  def create_jig_2(id=0, name="", type=0, capacity=0, jig_offset=p[0,0,0,0,0,0]):
      # iformation about used jigs
      return struct(id=id, name=name, type=type, capacity=capacity, jig_offset=jig_offset)
  end

  JIG2 = create_jig_2()
  JIGs = make_list(0, create_jig_2(), 20)

  JIGs.append(create_jig_2(id=1, name="3FG", type=1, capacity=1, jig_offset=p[0,0,0,0,0,0]))
  JIGs.append(create_jig_2(id=2, name="jig input", type=2, capacity=1, jig_offset=p[0,0,0,0,0,-3.927]))
  JIGs.append(create_jig_2(id=3, name="jig output", type=3, capacity=1, jig_offset=p[0,0,0,0,0,0.78]))
  JIGs.append(create_jig_2(id=6, name="jig bin", type=6, capacity=1, jig_offset=p[0,0,0,0,0,0]))
  JIGs.append(create_jig_2(id=7, name="jig sarstedt racks", type=7, capacity=1, jig_offset=p[0,0,-0.02,0,0,0]))
  JIGs.append(create_jig_2(id=8, name="NoK Bin", type=8, capacity=1, jig_offset=p[0,0,0,0,0,0]))
  JIGs.append(create_jig_2(id=9, name="Pick bott jig", type=9, capacity=1, jig_offset=p[0,0,0,0,0,0]))
  JIGs.append(create_jig_2(id=10, name="Place bott jig", type=10, capacity=1, jig_offset=p[0,0,0,0,0,0]))
  JIGs.append(create_jig_2(id=11, name="bottle shake jig", type=11, capacity=1, jig_offset=p[0,0,0,0,0,0]))
  JIGs.append(create_jig_2(id=12, name="Pick Vial jig", type=12, capacity=1, jig_offset=p[0,0,0,0,0,0]))
  JIGs.append(create_jig_2(id=13, name="Place Vial jig", type=13, capacity=1, jig_offset=p[0,0,0,0,0,0]))
  JIGs.append(create_jig_2(id=14, name="Liquid transfer jig", type=14, capacity=1, jig_offset=p[0,0,0,0,0,0]))
  JIGs.append(create_jig_2(id=15, name="Pick station jig", type=15, capacity=1, jig_offset=p[0,0,0,0,0,0]))
  JIGs.append(create_jig_2(id=16, name="Place station jig", type=16, capacity=1, jig_offset=p[0,0,0,0,0,0]))
  JIGs.append(create_jig_2(id=17, name="Weigh station jig", type=17, capacity=1, jig_offset=p[0,0,0,0,0,0]))
  JIGs.append(create_jig_2(id=18, name="Pick station 1", type=18, capacity=1, jig_offset=p[0,0,0,0,0,0]))
  JIGs.append(create_jig_2(id=19, name="Pick station 2", type=19, capacity=1, jig_offset=p[0,0,0,0,0,0]))
  JIGs.append(create_jig_2(id=20, name="Pick station 3", type=20, capacity=1, jig_offset=p[0,0,0,0,0,0]))
  $ 20 "Script: krish.script"
  def vibration_2():
  	set_analog_out(0,0.4)
  	sleep(0.6)
  	set_analog_out(0,0.0)
  	sleep(0.5)
  end

  def vibration_3():
  	set_analog_out(0,0.4)
  	sleep(0.3)
  	set_analog_out(0,0.0)
  	sleep(0.6)
  end

  def vibration_4():
  	set_analog_out(0,0.4)
  	sleep(0.25)
  	set_analog_out(0, 0.0)
  	sleep(1)
  end

  def vibration_1():
  	set_analog_out(0,0.4)
  	sleep(1)
  	set_analog_out(0,0.0)
  	sleep(0)
  end

  def move_tilt_in_steps(PowA_center, final_pose, steps):
  	i = 0
  	while i <= steps:
  		ratio = i / steps
  		pose_step = p[PowA_center[0] + ratio * (final_pose[0] - PowA_center[0]), PowA_center[1] + ratio * (final_pose[1] -PowA_center[1]),PowA_center[2] + ratio * (final_pose[2] - PowA_center[2]), PowA_center[3] + ratio * (final_pose[3] - PowA_center[3]), PowA_center[4] + ratio * (final_pose[4] - PowA_center[4]), PowA_center[5] + ratio * (final_pose[5] - PowA_center[5])]
  		movej(pose_step, a=1.2, v=0.15)
  		sleep(0.1)
  		i = i+1
  	end
  end

  def tilt_container(angle):
  	P_center = get_actual_tcp_pose()
  	hinge_offset = p[0,0,-0.23,0,0,0]
  	pivot_pose = pose_trans(P_center, hinge_offset)
  	pose_rel = pose_trans(pose_inv(pivot_pose), P_center)
  	angle_mid = (angle/2.0)*3.1416/180
  	angle_end = angle*3.1416/180
  	tilt_mid = p[0,0,0, -angle_mid, 0, 0]
  	tilt_end = p[0,0,0, -angle_end, 0, 0]
  	pose_rel_mid = pose_trans(tilt_mid, pose_rel)
  	pose_rel_end = pose_trans(tilt_end, pose_rel)
  	via_pose = pose_trans(pivot_pose, pose_rel_mid)
  	end_pose = pose_trans(pivot_pose, pose_rel_end)
  	movec(via_pose, end_pose, a=0.05, v=0.01, r=0.001)
  	P_center = get_actual_tcp_pose()
  end

  def scoop_powder(P_center):
  	#scoop_via_offset = p[0.05, 0.025, -0.03,0,0,0]
  	#scoop_end_offset = p[0.10, 0.05, -0.06, 0, 0,0]

  	#scoop_via_pose = pose_trans(scoop_start_pose, scoop_via_offset)
  	#scoop_end_pose = pose_trans(scoop_start_pose, scoop_end_offset)

  	#movel(scoop_start_pose, a=0.3, v=0.1)

  	#movec(scoop_via_pose, scoop_end_pose, a=0.3, v=0.1)

  	approach_offset = p[0.03,0,0.10,0,0,0]
  	scoop_radius = 0.03
  	#scoop_center = p[0, -0.01, 0.02, 0, 0, 1.5708]
  	tilt_down = p[0, 0, 0, -0.2618, 0, 0]
  	#scoop_out = p[0,0,0.10, 0, -0.2618,1.5708]
  	lift_offset = p[0, 0, 0.10, 0, 0, 0]
  	vibration_voltage = 4.0
  	vibration_time = 4.0

  	scoop_entry_pose = pose_trans(P_center, approach_offset)
  	movel(scoop_entry_pose, a=0.05, v=0.05)

  	scoop_start_rel = p[scoop_radius, 0, 0.02, 0, 0, 0]

  	rot_mid = p[0, 0, 0, 0, 0, 0.785]
  	rot_end = p[0, 0, 0, 0, 0, 1.5708]

  	scoop_via_rel = pose_trans(rot_mid, scoop_start_rel)
  	scoop_end_rel = pose_trans(rot_end, scoop_start_rel)

  	scoop_start_pose = pose_trans(P_center, scoop_start_rel)
  	scoop_via_pose = pose_trans(P_center, scoop_via_rel)
  	scoop_end_pose = pose_trans(P_center, scoop_end_rel)

  	movel(scoop_start_pose, a=0.03, v=0.05)

  	movec(scoop_via_pose, scoop_end_pose, a=0.03, v=0.05)

  	#scoop_center_pose = pose_trans(P_center, scoop_center)
  	#movel(scoop_center_pose, a=0.03, v=0.05)

  	tilted_pose = pose_trans(tilt_down, pose_trans(pose_inv(P_center), scoop_end_pose))
  	tilted_pose_in_base = pose_trans(P_center, tilted_pose)

  	movel(tilted_pose_in_base, a=0.03, v=0.05)

  	set_analog_out(0, vibration_voltage)
  	sleep(vibration_time)
  	set_analog_out(0, 0.0)

  	#scoop_out_pose = pose_trans(P_center, scoop_out)
  	#movel(scoop_out_pose, a=0.03, v=0.05)

  	tilt_pose_rel = pose_trans(pose_inv(P_center), tilted_pose_in_base)

  	lifted_pose_rel = pose_trans(lift_offset, tilt_pose_rel)

  	lifted_pose = pose_trans(P_center, lifted_pose_rel)
  	movel(lifted_pose, a=0.03, v=0.05)
  end
  $ 21 "Script: Weight_scale_socket.script"
  def get_weight():
  	socket_open("192.168.12.190", 3002)
  	textmsg("socket opened successfully!")
  	socket_send_string("GET_WEIGHT")
  	sync()
  	sleep(0.5)
  	receiveFromServ = socket_read_ascii_float(6)
  	while (receiveFromServ[0] <1):
  		sleep(0.5)
  		receiveFromServ = socket_read_ascii_float(1)
  		textmsg("retrying read:", receiveFromServ)
  	end
  	textmsg("Received weight:", receiveFromServ[1])
  	socket_close()
  	return receiveFromServ[1]
  end

  def tare_scale():
  	socket_open("192.168.12.190", 3002)
  	socket_send_string("TARE")
  	sleep(0.5)
  	socket_close()
  end

  def zero_scale():
  	socket_open("192.168.12.190", 3002)
  	socket_send_string("ZERO")
  	sleep(0.5)
  	socket_close()
  end
  $ 22 "BeforeStarts"
  $ 23 "uLM"
  $ 24 "CMD_Stop≔ False "
  global CMD_Stop=  False
  $ 25 "CMD_Abort≔ False "
  global CMD_Abort=  False
  $ 26 "CMD_Clear≔ False "
  global CMD_Clear=  False
  $ 27 "STATE≔1"
  global STATE=1
  $ 28 "STATE_Info≔''"
  global STATE_Info=""
  $ 29 "ARM_Referenced≔ False "
  global ARM_Referenced=  False
  $ 30 "zero_ftsensor()"
  zero_ftsensor()
  $ 31 "poses init"
  $ 32 "PSE_A≔p[0,0,0,0,0,0]"
  global PSE_A=p[0,0,0,0,0,0]
  $ 33 "PSE_A_H≔p[0,0,0,0,0,0]"
  global PSE_A_H=p[0,0,0,0,0,0]
  $ 34 "PSE_R≔p[0,0,0,0,0,0]"
  global PSE_R=p[0,0,0,0,0,0]
  $ 35 "PSE_R_H≔p[0,0,0,0,0,0]"
  global PSE_R_H=p[0,0,0,0,0,0]
  $ 36 "PSE_T≔p[0,0,0,0,0,0]"
  global PSE_T=p[0,0,0,0,0,0]
  $ 37 "PSE_T_H≔p[0,0,0,0,0,0]"
  global PSE_T_H=p[0,0,0,0,0,0]
  $ 38 "PSE_C_E≔p[0,0,0,0,0,0]"
  global PSE_C_E=p[0,0,0,0,0,0]
  $ 39 "PSE_C_H≔p[0,0,0,0,0,0]"
  global PSE_C_H=p[0,0,0,0,0,0]
  $ 40 "PSE_C_S≔p[0,0,0,0,0,0]"
  global PSE_C_S=p[0,0,0,0,0,0]
  $ 41 "init_home_by_cartesian_pose(p[0,-0.400,0.300,0,0,0])"
  init_home_by_cartesian_pose(p[0,-0.400,0.300,0,0,0])
  $ 42 "Clearing"
  $ 43 "reset_error()"
  reset_error()
  $ 44 "reset_warning()"
  reset_warning()
  $ 45 "uGo"
  $ 47 "ugo_init( True ,'http://192.168.12.120:10001')"
  ugo_init(  True  ,"http://192.168.12.120:10001")
  $ 48 "ugo_update_outputs()"
  ugo_update_outputs()
  $ 49 "App"
  $ 50 "'ADD APPLICATION SPECIFIC COMMANDS'"
  # 'ADD APPLICATION SPECIFIC COMMANDS'
  $ 51 "Tools"
  $ 52 "OBJ_Picked≔gripper_has_object()"
  global OBJ_Picked=gripper_has_object()
  $ 53 "If OBJ_Picked"
  if (OBJ_Picked):
    # begin: URCap Program Node
    #   Source: Robotiq_Grippers, 1.8.4.4844, Robotiq Inc.
    #   Type: Gripper Activate
    $ 54 "Gripper Activate"

    kill rq_gripper_communication_thread
    rq_gripper_communication_thread_started = False

    rq_init_comm_if_connected(9, "1")
    rq_init_comm_if_connected(2, "2")
    rq_init_comm_if_connected(3, "3")
    rq_init_comm_if_connected(4, "4")
    rq_print_connected_grippers()
    rq_gripper_communication_thread = run rq_gripper_communication()

    while(not rq_gripper_communication_thread_started):
        sync()
    end

    rq_set_max_current_for_all_grippers()

    reset_and_activate = False

    rq_activate_all_grippers(False)
    # end: URCap Program Node
  else:
    $ 55 "Else" "noBreak"
    # begin: URCap Program Node
    #   Source: Robotiq_Grippers, 1.8.4.4844, Robotiq Inc.
    #   Type: Gripper Activate
    $ 56 "Gripper Reset and Activate"

    kill rq_gripper_communication_thread
    rq_gripper_communication_thread_started = False

    rq_init_comm_if_connected(9, "1")
    rq_init_comm_if_connected(2, "2")
    rq_init_comm_if_connected(3, "3")
    rq_init_comm_if_connected(4, "4")
    rq_print_connected_grippers()
    rq_gripper_communication_thread = run rq_gripper_communication()

    while(not rq_gripper_communication_thread_started):
        sync()
    end

    rq_set_max_current_for_all_grippers()

    reset_and_activate = True

    rq_activate_all_grippers(True)
    # end: URCap Program Node
  end
  $ 57 "zero_ftsensor()"
  zero_ftsensor()
  $ 58 "EXTT"
  $ 59 "Set GRP_3F_Enable=Off"
  set_standard_digital_out(4, False)
  $ 60 "Set DO[6]=Off"
  set_standard_digital_out(6, False)
  $ 61 "Set GRP_3F_Decap=Off"
  set_standard_digital_out(3, False)
  $ 62 "Set GRP_3F_Cap=Off"
  set_standard_digital_out(2, False)
  $ 63 "Set GRP_3F_Open=Off"
  set_standard_digital_out(5, False)
  $ 64 "PSE_T≔get_tool_free_pose(dir=[0,0,0.150], move_in_base_frame=True)"
  global PSE_T=get_tool_free_pose(dir=[0,0,0.150], move_in_base_frame=True)
  $ 65 "If is_reachable(Base_const, [PSE_T])"
  if (is_reachable(p[0.0,0.0,0.0,0.0,0.0,0.0], [PSE_T])):
    $ 66 "MoveL"
    $ 67 "PSE_T" "breakAfter"
    movel(PSE_T, a=1.2, v=0.15)
  end
  $ 68 "powder dispensing variable init"
  $ 69 "Start_thread≔ False "
  global Start_thread=  False
  $ 70 "vib_mot_thread≔ False "
  global vib_mot_thread=  False
  $ 71 "kp≔0.00005"
  global kp=0.00005
  $ 72 "ki≔0.0005"
  global ki=0.0005
  $ 73 "kd≔0.002"
  global kd=0.002
  $ 74 "dt≔0.02"
  global dt=0.02
  $ 75 "Integral_error≔0"
  global Integral_error=0
  $ 76 "current_error≔0"
  global current_error=0
  $ 77 "previous_error≔0"
  global previous_error=0
  $ 78 "tilt_increment≔0"
  global tilt_increment=0
  $ 80 "diff≔0"
  global diff=0
  $ 81 "current_pose≔get_actual_tcp_pose()"
  global current_pose= get_actual_tcp_pose ()
  $ 82 "Relative_trans≔p[0.4902, -0.65024, -0.22623, 0.019, -0.263, -5.825]"
  global Relative_trans=p[0.4902, -0.65024, -0.22623, 0.019, -0.263, -5.825]
  $ 83 "ContA_plc_offst≔p[-0.00205, 0.02547, 0.03730, -0.03, -2.183, 6.165]"
  global ContA_plc_offst=p[-0.00205, 0.02547, 0.03730, -0.03, -2.183, 6.165]
  $ 84 "PowA_50_offset≔p[0.21808, -0.19943, 0.06584, 0, 0, 0]"
  global PowA_50_offset=p[0.21808, -0.19943, 0.06584, 0, 0, 0]
  $ 651 "Thread_1"
  thread Thread_1():
    while (True):
      $ 652 "If Start_thread≟ True "
      if (Start_thread ==   True  ):
        $ 653 "Weight_value≔get_weight()"
        global Weight_value=get_weight()
        $ 654 "sync()"
        sync()
      end
    end
  end
  threadId_Thread_1 = run Thread_1()
  $ 655 "Thread_2"
  thread Thread_2():
    while (True):
      $ 656 "Loop vib_mot_thread≟ True "
      thread Thread_while_656():
        while (True):
          $ 657 "diff≔Target_weight-Weight_value"
          global diff=Target_weight-Weight_value
          $ 658 "If diff>0.15"
          global thread_flag_658=0
          thread Thread_if_658():
            $ 660 "Set AO[0]=4.0"
            set_standard_analog_out(0, 0.4)
            thread_flag_658 = 1
          end
          if (diff>0.15):
            global thread_handler_658=run Thread_if_658()
            while (thread_flag_658 == 0):
              if not(diff>0.15):
                kill thread_handler_658
                thread_flag_658 = 2
              else:
                sync()
              end
            end
          else:
            thread_flag_658 = 2
          end
          if (thread_flag_658 == 2):
            $ 661 "ElseIf diff≥0.05 and diff≤0.15"
            global thread_flag_661=0
            thread Thread_if_661():
              $ 662 "vibration_2()"
              vibration_2()
              thread_flag_661 = 1
            end
            if (diff >= 0.05 and diff <= 0.15):
              global thread_handler_661=run Thread_if_661()
              while (thread_flag_661 == 0):
                if not(diff >= 0.05 and diff <= 0.15):
                  kill thread_handler_661
                  thread_flag_661 = 2
                else:
                  sync()
                end
              end
            else:
              thread_flag_661 = 2
            end
            if (thread_flag_661 == 2):
              $ 663 "ElseIf diff≥0.01 and diff<0.05"
              if (diff >= 0.01 and diff<0.05):
                $ 664 "vibration_3()"
                vibration_3()
              else:
                $ 665 "ElseIf diff>0 and diff<0.01"
                if (diff>0 and diff<0.01):
                  $ 666 "vibration_4()"
                  vibration_4()
                else:
                  $ 667 "Else" "noBreak"
                  $ 668 "Set AO[0]=0.0"
                  set_standard_analog_out(0, 0.0)
                end
              end
            end
          end
        end
      end
      if (vib_mot_thread ==   True  ):
        global thread_handler_656=run Thread_while_656()
        while (vib_mot_thread ==   True  ):
          sync()
        end
        kill thread_handler_656
      end
      $ 671 "sync()"
      sync()
    end
  end
  threadId_Thread_2 = run Thread_2()
  while (True):
    $ 85 "Robot Program"
    $ 86 "MAIN"
    $ 87 "command_manager(external_control='uGO', cond_suspend=(ITM_Manipulated and AMR_AtTarget and AMR_Charging and AMR_Battery<40), cond_unsuspend=(AMR_Battery≟60))"
    command_manager(external_control="uGO", cond_suspend=(ITM_Manipulated  and  AMR_AtTarget  and  AMR_Charging  and  AMR_Battery<40), cond_unsuspend=(AMR_Battery == 60))
    $ 88 "log_state(STATE_Info)"
    log_state(STATE_Info)
    $ 89 "Switch STATE"
    switch_1 = STATE
    $ 90 "Case 1"
    if (1 == switch_1):
      $ 91 "Stopping"
      $ 92 "STATE_Info≔'Stopping'"
      global STATE_Info="Stopping"
      $ 93 "end_freedrive_mode()"
      end_freedrive_mode()
      $ 94 "Set"
      set_tcp(p[0.0,0.0,0.161,3.1415,0.0,0.0])
      $ 95 "PSE_T≔get_tool_free_pose(dir=[0,0,0.150], move_in_base_frame=True)"
      global PSE_T=get_tool_free_pose(dir=[0,0,0.150], move_in_base_frame=True)
      $ 96 "If is_reachable(Base_const, [PSE_T])"
      if (is_reachable(p[0.0,0.0,0.0,0.0,0.0,0.0], [PSE_T])):
        $ 97 "MoveL"
        $ 98 "PSE_T" "breakAfter"
        movel(PSE_T, a=1.2, v=0.15)
      end
      $ 99 "do_transition(keep_rxry=OBJ_Picked, r=0)"
      do_transition(keep_rxry=OBJ_Picked, r=0)
      $ 108 "Call Sub_AMR_MiR_V3"
      Sub_AMR_MiR_V3()
      $ 109 "If stopping() and AMR_Done"
      if (stopping()  and  AMR_Done):
        $ 110 "STATE≔2"
        global STATE=2
        $ 111 "ugo_update_outputs()"
        ugo_update_outputs()
      end
    elif (2 == switch_1):
      $ 112 "Case 2"
      $ 113 "Stopped"
      $ 114 "STATE_Info≔'Stopped'"
      global STATE_Info="Stopped"
      $ 115 "Call Sub_AMR_MiR_V3"
      Sub_AMR_MiR_V3()
      $ 116 "If CMD_Reset"
      if (CMD_Reset):
        $ 117 "STATE≔3"
        global STATE=3
        $ 118 "ugo_update_outputs()"
        ugo_update_outputs()
      end
    elif (3 == switch_1):
      $ 119 "Case 3"
      $ 120 " Resetting"
      $ 121 "STATE_Info≔'Resetting'"
      global STATE_Info="Resetting"
      $ 122 "uML"
      $ 123 "reset_error()"
      reset_error()
      $ 124 "reset_warning()"
      reset_warning()
      $ 125 "PROCESS_Step≔0"
      global PROCESS_Step=0
      $ 126 "PROCESS_Info≔''"
      global PROCESS_Info=""
      $ 127 "ARM_Referenced≔ False "
      global ARM_Referenced=  False
      $ 128 "WRK_Done≔ False "
      global WRK_Done=  False
      $ 129 "ITM_Prepared≔ False "
      global ITM_Prepared=  False
      $ 130 "ITM_Manipulated≔ False "
      global ITM_Manipulated=  False
      $ 131 "STP≔0"
      global STP=0
      $ 132 "Action≔0"
      global Action=0
      $ 133 "Action_Info≔''"
      global Action_Info=""
      $ 134 "ITM_ID≔0"
      global ITM_ID=0
      $ 135 "JIG≔0"
      global JIG=0
      $ 136 "JIG_Slot≔0"
      global JIG_Slot=0
      $ 137 "Task_info≔''"
      global Task_info=""
      $ 138 "Set"
      set_tcp(p[0.0,0.0,0.161,3.1415,0.0,0.0])
      $ 139 "App"
      $ 140 "'ADD APPLICATION SPECIFIC COMMANDS'"
      # 'ADD APPLICATION SPECIFIC COMMANDS'
      $ 141 "OBJ_Type≔0"
      global OBJ_Type=0
      $ 142 "OBJ_Nbr≔0"
      global OBJ_Nbr=0
      $ 143 "If CNT_Rack_Output≥50"
      if (CNT_Rack_Output >= 50):
        $ 144 "CNT_Rack_Output≔0"
        global CNT_Rack_Output=0
      end
      $ 145 "TASK≔struct(ID=0, NAVI=struct(target=0, footprint=0, protectiveOff=0, dock=0), WORK=struct(ITM_ID_Src=0, JIG_ID_Src=0, OBJ_Nbr_Src=0, ACT_Src=0, ITM_ID_Tgt=0, JIG_ID_Tgt=0, OBJ_Nbr_Tgt=0, ACT_Tgt=0, OBJ_Type=0))"
      global TASK=struct(ID=0, NAVI=struct(target=0, footprint=0, protectiveOff=0, dock=0), WORK=struct(ITM_ID_Src=0, JIG_ID_Src=0, OBJ_Nbr_Src=0, ACT_Src=0, ITM_ID_Tgt=0, JIG_ID_Tgt=0, OBJ_Nbr_Tgt=0, ACT_Tgt=0, OBJ_Type=0))
      $ 146 "Call Sub_AMR_MiR_V3"
      Sub_AMR_MiR_V3()
      $ 147 "If resetting() and AMR_Done"
      if (resetting()  and  AMR_Done):
        $ 148 "STATE≔4"
        global STATE=4
        $ 149 "ugo_update_outputs()"
        ugo_update_outputs()
      end
    elif (4 == switch_1):
      $ 150 "Case 4"
      $ 151 "Idle"
      $ 152 "STATE_Info≔'Idle'"
      global STATE_Info="Idle"
      $ 153 "If CMD_Start"
      if (CMD_Start):
        $ 154 "STATE≔5"
        global STATE=5
        $ 155 "ugo_update_outputs()"
        ugo_update_outputs()
      end
    elif (5 == switch_1):
      $ 156 "Case 5"
      $ 157 "Starting"
      $ 158 "STATE_Info≔'Starting'"
      global STATE_Info="Starting"
      $ 159 "'ADD COMMANDS WHAT TO START WITH'"
      # 'ADD COMMANDS WHAT TO START WITH'
      $ 160 "Call Sub_AMR_MiR_V3"
      Sub_AMR_MiR_V3()
      $ 161 "get ugo data"
      $ 162 "Assign Tasks"
      $ 163 "TASK.ID = ugo_get_task()"
      TASK.ID = ugo_get_task()
      $ 164 "If TASK.ID≟1"
      if (TASK.ID == 1):
        $ 165 "Task_info≔'Charge'"
        global Task_info="Charge"
        $ 166 "Parameters"
        $ 167 "AMR_PosTarget≔1"
        global AMR_PosTarget=1
      else:
        $ 168 "ElseIf TASK.ID≟9"
        if (TASK.ID == 9):
          $ 169 "'Pick Sarstedt Rack from Variable source'"
          # 'Pick Sarstedt Rack from Variable source'
          $ 170 "Task_info≔'Navigate to Target'"
          global Task_info="Navigate to Target"
          $ 171 "Parameters"
          $ 172 "AMR_PosTarget≔UGO.read_input('00','ITM_ID')"
          global AMR_PosTarget=UGO.read_input("00","ITM_ID")
        else:
          $ 173 "ElseIf TASK.ID≟99"
          if (TASK.ID == 99):
            $ 174 "Task_info≔'Pick rack pipet'"
            global Task_info="Pick rack pipet"
            $ 175 "Parameters"
            $ 176 "ITM_ID≔1"
            global ITM_ID=1
            $ 177 "OBJ_Type≔9"
            global OBJ_Type=9
            $ 178 "JIG≔18"
            global JIG=18
            $ 179 "AMR_PosTarget≔3"
            global AMR_PosTarget=3
          else:
            $ 180 "ElseIf TASK.ID≟98"
            if (TASK.ID == 98):
              $ 181 "Task_info≔'Place rack pipet'"
              global Task_info="Place rack pipet"
              $ 182 "Parameters"
              $ 183 "ITM_ID≔1"
              global ITM_ID=1
              $ 184 "OBJ_Type≔9"
              global OBJ_Type=9
              $ 185 "JIG≔19"
              global JIG=19
              $ 186 "AMR_PosTarget≔2"
              global AMR_PosTarget=2
            else:
              $ 187 "Else" "noBreak"
              $ 188 "set_error(ERROR_WRONG_ORDER)"
              set_error(ERROR_WRONG_ORDER)
            end
          end
        end
      end
      $ 189 "test ugo"
      $ 190 "Wait: 0.2"
      sleep(0.2)
      $ 191 "ugo_update_outputs()"
      ugo_update_outputs()
      $ 192 "If starting() and AMR_Done"
      if (starting()  and  AMR_Done):
        $ 193 "log_message(Task_info, 'New Task: ')"
        log_message(Task_info, "New Task: ")
        $ 194 "log_message(to_str(TASK.ID), 'Task_ID: ')"
        log_message(to_str(TASK.ID), "Task_ID: ")
        $ 195 "do_transition(keep_rxry=OBJ_Picked)"
        do_transition(keep_rxry=OBJ_Picked)
        $ 196 "STATE≔6"
        global STATE=6
        $ 197 "ugo_update_outputs()"
        ugo_update_outputs()
      end
    elif (6 == switch_1):
      $ 198 "Case 6"
      $ 199 "Execute"
      $ 200 "STATE_Info≔'Execute'"
      global STATE_Info="Execute"
      $ 201 "If  not CMD_Hold and not CMD_Suspend"
      global thread_flag_201=0
      thread Thread_if_201():
        $ 202 "Switch PROCESS_Step"
        switch_2 = PROCESS_Step
        $ 203 "Case 0"
        if (0 == switch_2):
          $ 204 "PROCESS_Info≔'process control'"
          global PROCESS_Info="process control"
          $ 205 "log_process(PROCESS_Info)"
          log_process(PROCESS_Info)
          $ 206 "process control"
          $ 207 "If  not AMR_AtTarget"
          if (  not  AMR_AtTarget):
            $ 208 "PROCESS_Step≔1"
            global PROCESS_Step=1
          else:
            $ 209 "ElseIf (( not ITM_Prepared and  not WRK_Done) or (ITM_Prepared and WRK_Done))"
            if (((  not  ITM_Prepared  and    not  WRK_Done)  or  (ITM_Prepared  and  WRK_Done))):
              $ 210 "PROCESS_Step≔2"
              global PROCESS_Step=2
            else:
              $ 211 "ElseIf  not WRK_Done"
              if (  not  WRK_Done):
                $ 212 "PROCESS_Step≔3"
                global PROCESS_Step=3
              else:
                $ 213 "Else" "noBreak"
                $ 214 "task finished"
                $ 215 "PROCESS_Info≔''"
                global PROCESS_Info=""
                $ 216 "STATE≔7"
                global STATE=7
                $ 217 "ugo_update_outputs()"
                ugo_update_outputs()
              end
            end
          end
        elif (1 == switch_2):
          $ 218 "Case 1"
          $ 219 "navigate"
          $ 220 "'MOVING THE uML'"
          # 'MOVING THE uML'
          $ 221 "PROCESS_Info≔'move to target'"
          global PROCESS_Info="move to target"
          $ 222 "log_process(PROCESS_Info)"
          log_process(PROCESS_Info)
          $ 223 "If TASK.ID≟1"
          if (TASK.ID == 1):
            $ 224 "Action≔51"
            global Action=51
          else:
            $ 225 "Else" "noBreak"
            $ 226 "Action≔52"
            global Action=52
          end
          $ 227 "Call Sub_AMR_MiR_V3"
          Sub_AMR_MiR_V3()
          $ 228 "If AMR_Done"
          if (AMR_Done):
            $ 229 "PROCESS_Step≔0"
            global PROCESS_Step=0
          end
        elif (2 == switch_2):
          $ 230 "Case 2"
          $ 231 "prepare"
          $ 232 "'THINGS THAT HAVE TO BE DONE ONCE IN A SEQUENCE,WORKFLOW'"
          # 'THINGS THAT HAVE TO BE DONE ONCE IN A SEQUENCE,WORKFLOW'
          $ 233 "PROCESS_Info≔'prepare for work'"
          global PROCESS_Info="prepare for work"
          $ 234 "log_process(PROCESS_Info)"
          log_process(PROCESS_Info)
          $ 235 "If TASK.WORK.ITM_ID_Src>1"
          if (TASK.WORK.ITM_ID_Src>1):
            $ 236 "ITM_ID≔TASK.WORK.ITM_ID_Src"
            global ITM_ID=TASK.WORK.ITM_ID_Src
          else:
            $ 237 "ElseIf TASK.WORK.ITM_ID_Tgt>1"
            if (TASK.WORK.ITM_ID_Tgt>1):
              $ 238 "ITM_ID≔TASK.WORK.ITM_ID_Tgt"
              global ITM_ID=TASK.WORK.ITM_ID_Tgt
            end
          end
          $ 239 "If  not ARM_Referenced and (ITM_ID≠0)"
          if (  not  ARM_Referenced  and  (ITM_ID != 0)):
            $ 240 "STP≔1"
            global STP=1
          else:
            $ 241 "ElseIf ARM_Referenced or (ITM_ID≟0)"
            if (ARM_Referenced  or  (ITM_ID == 0)):
              $ 242 "STP≔2"
              global STP=2
            end
          end
          $ 243 "Switch STP"
          switch_3 = STP
          $ 244 "Case 1"
          if (1 == switch_3):
            $ 245 "reference"
            $ 246 "STP_Info≔'reference at target position'"
            global STP_Info="reference at target position"
            $ 247 "log_step(STP_Info)"
            log_step(STP_Info)
            $ 248 "If ITM_ID≟1"
            if (ITM_ID == 1):
              $ 249 "CAM_Done≔ True "
              global CAM_Done=  True
            else:
              $ 250 "Else" "noBreak"
              $ 251 "Action≔131"
              global Action=131
              $ 252 "Call Sub_Vision_V18"
              Sub_Vision_V18()
            end
            $ 254 "If CAM_Done and  not ERROR.FLAG"
            if (CAM_Done  and    not  ERROR.FLAG):
              $ 255 "log_step('ARM referenced')"
              log_step("ARM referenced")
              $ 256 "ARM_Referenced≔ True "
              global ARM_Referenced=  True
            end
          elif (2 == switch_3):
            $ 257 "Case 2"
            $ 258 "manipulate"
            $ 259 "STP_Info≔'manipulate item'"
            global STP_Info="manipulate item"
            $ 260 "log_step(STP_Info)"
            log_step(STP_Info)
            $ 261 "'In case pressing button is needed'"
            # 'In case pressing button is needed'
            $ 262 "If found_in_list(ITM_ID, ITM_ID_List)"
            if (found_in_list(ITM_ID, ITM_ID_List)):
              $ 263 "Switch ITM_ID"
              switch_4 = ITM_ID
              $ 264 "Case 0"
              if (0 == switch_4):
                $ 265 "ITM_Manipulated≔ not ITM_Manipulated"
                global ITM_Manipulated=  not  ITM_Manipulated
              elif (1 == switch_4):
                $ 266 "Case 1"
                $ 267 "ITM_Manipulated≔ not ITM_Manipulated"
                global ITM_Manipulated=  not  ITM_Manipulated
              elif (2 == switch_4):
                $ 268 "Case 2"
              else:
                $ 278 "Default Case"
                $ 279 "ITM_Manipulated≔ not ITM_Manipulated"
                global ITM_Manipulated=  not  ITM_Manipulated
              end
            end
          end
          $ 280 "ITM_Prepared≔(ITM_Manipulated or  not found_in_list(ITM_ID, ITM_ID_List)) and (ARM_Referenced or ITM_ID≟0) and  not WRK_Done"
          global ITM_Prepared=(ITM_Manipulated  or    not  found_in_list(ITM_ID, ITM_ID_List))  and  (ARM_Referenced  or  ITM_ID == 0)  and    not  WRK_Done
          $ 281 "STP≔0"
          global STP=0
          $ 282 "STP_Info≔''"
          global STP_Info=""
          $ 283 "PROCESS_Step≔0"
          global PROCESS_Step=0
        elif (3 == switch_2):
          $ 284 "Case 3"
          $ 285 "work"
          $ 286 "'ADD EVERY MACHINE, OBJECT, STATION TO WORK ON'"
          # 'ADD EVERY MACHINE, OBJECT, STATION TO WORK ON'
          $ 287 "Switch ITM_ID"
          switch_3 = ITM_ID
          $ 288 "Case 1"
          if (1 == switch_3):
            $ 289 "uLM"
            $ 290 "If TASK.ID≟12"
            if (TASK.ID == 12):
              $ 291 "fill racks"
              $ 292 "Action≔151"
              global Action=151
              $ 293 "Call Sub_Vision_V18"
              Sub_Vision_V18()
              $ 294 "If  not ERROR.FLAG"
              if (  not  ERROR.FLAG):
                $ 295 "Actions for the task"
                $ 296 "Action≔1"
                global Action=1
                $ 297 "JIG≔2"
                global JIG=2
                $ 298 "JIG_Slot≔CAM_Result[0]"
                global JIG_Slot=CAM_Result[0]
                $ 299 "OBJ_Nbr≔CAM_Result[0]"
                global OBJ_Nbr=CAM_Result[0]
                $ 300 "OBJ_Type≔2"
                global OBJ_Type=2
                $ 301 "Call Sub_Action_V4"
                Sub_Action_V4()
                $ 302 "If OBJ_Picked"
                if (OBJ_Picked):
                  $ 303 "CAM_Result.remove(0)"
                  CAM_Result.remove(0)
                  $ 304 "PRC_TubCounter≔PRC_TubCounter+1"
                  global PRC_TubCounter=PRC_TubCounter+1
                  $ 305 "If PRC_TubCounter%4≟0"
                  if (PRC_TubCounter%4 == 0):
                    $ 306 "JIG_Slot≔4"
                    global JIG_Slot=4
                  else:
                    $ 307 "Else" "noBreak"
                    $ 308 "JIG_Slot≔PRC_TubCounter%4"
                    global JIG_Slot=PRC_TubCounter%4
                  end
                  $ 309 "OBJ_Nbr≔ceil(PRC_TubCounter/4)"
                  global OBJ_Nbr=ceil(PRC_TubCounter/4)
                  $ 310 "Action≔2"
                  global Action=2
                  $ 311 "JIG≔4"
                  global JIG=4
                  $ 312 "Call Sub_Action_V4"
                  Sub_Action_V4()
                  $ 313 "Action≔151"
                  global Action=151
                  $ 314 "Call Sub_Vision_V18"
                  Sub_Vision_V18()
                end
              end
              $ 315 "If (CAM_Captures≥CAM_PRM_Retries) or (PRC_TubCounter≥32)"
              if ((CAM_Captures >= CAM_PRM_Retries)  or  (PRC_TubCounter >= 32)):
                $ 316 "PROCESS_Step≔0"
                global PROCESS_Step=0
                $ 317 "WRK_Done≔ True "
                global WRK_Done=  True
              end
            else:
              $ 318 "ElseIf TASK.ID≟49"
              if (TASK.ID == 49):
                $ 319 "Pick Powder container"
                $ 320 "Action≔131"
                global Action=131
                $ 321 "Call Sub_Vision_V18"
                Sub_Vision_V18()
                $ 322 "Action≔35"
                global Action=35
                $ 323 "Call Sub_Action_V4"
                Sub_Action_V4()
                $ 324 "PROCESS_Step≔0"
                global PROCESS_Step=0
                $ 325 "WRK_Done≔ True "
                global WRK_Done=  True
              else:
                $ 326 "ElseIf TASK.ID≟50"
                if (TASK.ID == 50):
                  $ 327 "Decap containers"
                  $ 328 "Action≔36"
                  global Action=36
                  $ 329 "Call Sub_Action_V4"
                  Sub_Action_V4()
                  $ 330 "PROCESS_Step≔0"
                  global PROCESS_Step=0
                  $ 331 "WRK_Done≔ True "
                  global WRK_Done=  True
                else:
                  $ 332 "ElseIf TASK.ID≟51"
                  if (TASK.ID == 51):
                    $ 333 "Detect Spatula and transfer powder"
                    $ 334 "Action≔131"
                    global Action=131
                    $ 335 "Call Sub_Vision_V18"
                    Sub_Vision_V18()
                    $ 336 "Action≔37"
                    global Action=37
                    $ 337 "Call Sub_Action_V4"
                    Sub_Action_V4()
                    $ 338 "PROCESS_Step≔0"
                    global PROCESS_Step=0
                    $ 339 "WRK_Done≔ True "
                    global WRK_Done=  True
                  else:
                    $ 340 "ElseIf TASK.ID≟52"
                    if (TASK.ID == 52):
                      $ 341 "Pick PowderA container"
                      $ 342 "Action≔131"
                      global Action=131
                      $ 343 "Call Sub_Vision_V18"
                      Sub_Vision_V18()
                      $ 344 "Action≔38"
                      global Action=38
                      $ 345 "Call Sub_Action_V4"
                      Sub_Action_V4()
                      $ 346 "PROCESS_Step≔0"
                      global PROCESS_Step=0
                      $ 347 "WRK_Done≔ True "
                      global WRK_Done=  True
                    else:
                      $ 348 "ElseIf TASK.ID≟53"
                      if (TASK.ID == 53):
                        $ 349 "Decap containerA"
                        $ 350 "Action≔39"
                        global Action=39
                        $ 351 "Call Sub_Action_V4"
                        Sub_Action_V4()
                        $ 352 "PROCESS_Step≔0"
                        global PROCESS_Step=0
                        $ 353 "WRK_Done≔ True "
                        global WRK_Done=  True
                      else:
                        $ 354 "ElseIf TASK.ID≟54"
                        if (TASK.ID == 54):
                          $ 355 "Dispense PowderA"
                          $ 356 "Action≔131"
                          global Action=131
                          $ 357 "Call Sub_Vision_V18"
                          Sub_Vision_V18()
                          $ 358 "Action≔40"
                          global Action=40
                          $ 359 "Call Sub_Action_V4"
                          Sub_Action_V4()
                          $ 360 "PROCESS_Step≔0"
                          global PROCESS_Step=0
                          $ 361 "WRK_Done≔ True "
                          global WRK_Done=  True
                        else:
                          $ 362 "ElseIf TASK.ID≟54"
                          if (TASK.ID == 54):
                            $ 363 "Dispense PowderA"
                            $ 364 "Action≔131"
                            global Action=131
                            $ 365 "Call Sub_Vision_V18"
                            Sub_Vision_V18()
                            $ 366 "Action≔40"
                            global Action=40
                            $ 367 "Call Sub_Action_V4"
                            Sub_Action_V4()
                            $ 368 "PROCESS_Step≔0"
                            global PROCESS_Step=0
                            $ 369 "WRK_Done≔ True "
                            global WRK_Done=  True
                          else:
                            $ 370 "ElseIf TASK.ID≟99"
                            if (TASK.ID == 99):
                              $ 371 "Pick rack pipet"
                              $ 372 "Action≔131"
                              global Action=131
                              $ 373 "Call Sub_Vision_V18"
                              Sub_Vision_V18()
                              $ 374 "Action≔5"
                              global Action=5
                              $ 375 "Call Sub_Action_V4"
                              Sub_Action_V4()
                              $ 376 "PROCESS_Step≔0"
                              global PROCESS_Step=0
                              $ 377 "WRK_Done≔ True "
                              global WRK_Done=  True
                            else:
                              $ 378 "ElseIf TASK.ID≟98"
                              if (TASK.ID == 98):
                                $ 379 "Pick rack pipet"
                                $ 380 "Action≔131"
                                global Action=131
                                $ 381 "Call Sub_Vision_V18"
                                Sub_Vision_V18()
                                $ 382 "Action≔6"
                                global Action=6
                                $ 383 "Call Sub_Action_V4"
                                Sub_Action_V4()
                                $ 384 "PROCESS_Step≔0"
                                global PROCESS_Step=0
                                $ 385 "WRK_Done≔ True "
                                global WRK_Done=  True
                              end
                            end
                          end
                        end
                      end
                    end
                  end
                end
              end
            end
          elif (2 == switch_3):
            $ 386 "Case 2"
          elif (5 == switch_3):
            $ 428 "Case 5"
          elif (20 == switch_3):
            $ 436 "Case 20"
          elif (43 == switch_3):
            $ 498 "Case 43"
          else:
            $ 506 "Default Case"
            $ 507 "WRK_Done≔ True "
            global WRK_Done=  True
            $ 508 "PROCESS_Step≔0"
            global PROCESS_Step=0
          end
        end
        thread_flag_201 = 1
      end
      if (  not  CMD_Hold and not CMD_Suspend):
        global thread_handler_201=run Thread_if_201()
        while (thread_flag_201 == 0):
          if not(  not  CMD_Hold and not CMD_Suspend):
            kill thread_handler_201
            thread_flag_201 = 2
          else:
            sync()
          end
        end
      else:
        thread_flag_201 = 2
      end
      $ 509 "If CMD_Hold"
      if (CMD_Hold):
        $ 510 "STATE≔9"
        global STATE=9
        $ 511 "ugo_update_outputs()"
        ugo_update_outputs()
      else:
        $ 512 "ElseIf CMD_Suspend"
        if (CMD_Suspend):
          $ 513 "STATE≔12"
          global STATE=12
          $ 514 "ugo_update_outputs()"
          ugo_update_outputs()
        end
      end
    elif (7 == switch_1):
      $ 515 "Case 7"
      $ 516 "Completing"
      $ 517 "STATE_Info≔'Completing'"
      global STATE_Info="Completing"
      $ 518 "'ADD COMMANDS FOR COMPLETING THE PROCESS'"
      # 'ADD COMMANDS FOR COMPLETING THE PROCESS'
      $ 519 "do_transition(keep_rxry=OBJ_Picked)"
      do_transition(keep_rxry=OBJ_Picked)
      $ 520 "Call Sub_AMR_MiR_V3"
      Sub_AMR_MiR_V3()
      $ 521 "If completing() and AMR_Done"
      if (completing()  and  AMR_Done):
        $ 522 "STATE≔8"
        global STATE=8
        $ 523 "ugo_update_outputs()"
        ugo_update_outputs()
      end
    elif (8 == switch_1):
      $ 524 "Case 8"
      $ 525 "Complete"
      $ 526 "STATE_Info≔'Complete'"
      global STATE_Info="Complete"
      $ 527 "If CMD_Reset"
      if (CMD_Reset):
        $ 528 "STATE≔3"
        global STATE=3
        $ 529 "ugo_update_outputs()"
        ugo_update_outputs()
      end
    elif (9 == switch_1):
      $ 530 "Case 9"
      $ 531 "Holding"
      $ 532 "STATE_Info≔'Holding'"
      global STATE_Info="Holding"
      $ 533 "stopl(0.5)"
      stopl(0.5)
      $ 534 "Call Sub_AMR_MiR_V3"
      Sub_AMR_MiR_V3()
      $ 535 "If holding() and AMR_Done"
      if (holding()  and  AMR_Done):
        $ 536 "STATE≔10"
        global STATE=10
        $ 537 "ugo_update_outputs()"
        ugo_update_outputs()
      end
    elif (10 == switch_1):
      $ 538 "Case 10"
      $ 539 "Held"
      $ 540 "STATE_Info≔'Held'"
      global STATE_Info="Held"
      $ 541 "If CMD_Unhold"
      if (CMD_Unhold):
        $ 542 "end_freedrive_mode()"
        end_freedrive_mode()
        $ 543 "STATE≔11"
        global STATE=11
        $ 544 "ugo_update_outputs()"
        ugo_update_outputs()
      else:
        $ 545 "ElseIf FNC_Freedrive"
        if (FNC_Freedrive):
          $ 546 "freedrive_mode()"
          freedrive_mode()
        else:
          $ 547 "Else" "noBreak"
          $ 548 "end_freedrive_mode()"
          end_freedrive_mode()
        end
      end
    elif (11 == switch_1):
      $ 549 "Case 11"
      $ 550 "Unholding"
      $ 551 "STATE_Info≔'Unholding'"
      global STATE_Info="Unholding"
      $ 552 "Clearing"
      $ 553 "Switch ERROR.ID"
      switch_2 = ERROR.ID
      $ 554 "Case 1002"
      if (1002 == switch_2):
        $ 555 "AMR_AtTarget≔ False "
        global AMR_AtTarget=  False
        $ 556 "ARM_Referenced≔ False "
        global ARM_Referenced=  False
        $ 557 "ITM_Prepared≔ False "
        global ITM_Prepared=  False
        $ 558 "PROCESS_Step≔1"
        global PROCESS_Step=1
      elif (2007 == switch_2):
        $ 559 "Case 2007"
        $ 560 "PROCESS_Step≔1"
        global PROCESS_Step=1
      end
      $ 561 "reset_error()"
      reset_error()
      $ 562 "reset_warning()"
      reset_warning()
      $ 563 "OBJ_Picked≔gripper_has_object()"
      global OBJ_Picked=gripper_has_object()
      $ 564 "Call Sub_AMR_MiR_V3"
      Sub_AMR_MiR_V3()
      $ 565 "If unholding() and AMR_Done"
      if (unholding()  and  AMR_Done):
        $ 566 "STATE≔6"
        global STATE=6
        $ 567 "ugo_update_outputs()"
        ugo_update_outputs()
      end
    elif (12 == switch_1):
      $ 568 "Case 12"
      $ 569 "Suspending"
      $ 570 "STATE_Info≔'Suspending'"
      global STATE_Info="Suspending"
      $ 571 "PROCESS_Info≔str_cat(PROCESS_Info, ' suspended')"
      global PROCESS_Info=str_cat(PROCESS_Info, " suspended")
      $ 572 "If suspending()"
      if (suspending()):
        $ 573 "STATE≔13"
        global STATE=13
        $ 574 "ugo_update_outputs()"
        ugo_update_outputs()
      end
    elif (13 == switch_1):
      $ 575 "Case 13"
      $ 576 "Suspended"
      $ 577 "STATE_Info≔'Suspended'"
      global STATE_Info="Suspended"
      $ 578 "Call Sub_AMR_MiR_V3"
      Sub_AMR_MiR_V3()
      $ 579 "If CMD_Unsuspend"
      if (CMD_Unsuspend):
        $ 580 "STATE≔14"
        global STATE=14
        $ 581 "ugo_update_outputs()"
        ugo_update_outputs()
      end
    elif (14 == switch_1):
      $ 582 "Case 14"
      $ 583 "Unsuspending"
      $ 584 "STATE_Info≔'Unsuspending'"
      global STATE_Info="Unsuspending"
      $ 585 "PROCESS_Step≔0"
      global PROCESS_Step=0
      $ 586 "If unsuspending()"
      if (unsuspending()):
        $ 587 "STATE≔6"
        global STATE=6
        $ 588 "ugo_update_outputs()"
        ugo_update_outputs()
      end
    elif (15 == switch_1):
      $ 589 "Case 15"
      $ 590 "Aborting"
      $ 591 "STATE_Info≔'Aborting'"
      global STATE_Info="Aborting"
      $ 592 "If aborting()"
      if (aborting()):
        $ 593 "STATE≔16"
        global STATE=16
        $ 594 "ugo_update_outputs()"
        ugo_update_outputs()
      end
    elif (16 == switch_1):
      $ 595 "Case 16"
      $ 596 "Aborted"
      $ 597 "STATE_Info≔'Aborted'"
      global STATE_Info="Aborted"
      $ 598 "If CMD_Clear"
      if (CMD_Clear):
        $ 599 "STATE≔17"
        global STATE=17
        $ 600 "ugo_update_outputs()"
        ugo_update_outputs()
      end
    elif (17 == switch_1):
      $ 601 "Case 17"
      $ 602 "Clearing"
      $ 603 "STATE_Info≔'Clearing'"
      global STATE_Info="Clearing"
      $ 604 "Clearing"
      $ 605 "reset_warning()"
      reset_warning()
      $ 606 "reset_error()"
      reset_error()
      $ 607 "If clearing()"
      if (clearing()):
        $ 608 "STATE≔2"
        global STATE=2
        $ 609 "ugo_update_outputs()"
        ugo_update_outputs()
      end
    end
    $ 610 "log_state(STATE_Info)"
    log_state(STATE_Info)
    $ 611 "log_warning(WARNING.MSG)"
    log_warning(WARNING.MSG)
    $ 612 "log_error(ERROR.MSG)"
    log_error(ERROR.MSG)
    $ 613 "Times"
    $ 614 "Switch STATE"
    switch_1 = STATE
    $ 615 "Case 1"
    if (1 == switch_1):
      $ 616 "TM_St_Stopping≔get_time(STATE_Times[STATE-1])"
      global TM_St_Stopping=get_time(STATE_Times[STATE-1])
    elif (2 == switch_1):
      $ 617 "Case 2"
      $ 618 "TM_St_Stopped≔get_time(STATE_Times[STATE-1])"
      global TM_St_Stopped=get_time(STATE_Times[STATE-1])
    elif (3 == switch_1):
      $ 619 "Case 3"
      $ 620 "TM_St_Resetting≔get_time(STATE_Times[STATE-1])"
      global TM_St_Resetting=get_time(STATE_Times[STATE-1])
    elif (4 == switch_1):
      $ 621 "Case 4"
      $ 622 "TM_St_Idle≔get_time(STATE_Times[STATE-1])"
      global TM_St_Idle=get_time(STATE_Times[STATE-1])
    elif (5 == switch_1):
      $ 623 "Case 5"
      $ 624 "TM_St_Starting≔get_time(STATE_Times[STATE-1])"
      global TM_St_Starting=get_time(STATE_Times[STATE-1])
    elif (6 == switch_1):
      $ 625 "Case 6"
      $ 626 "TM_St_Execute≔get_time(STATE_Times[STATE-1])"
      global TM_St_Execute=get_time(STATE_Times[STATE-1])
    elif (7 == switch_1):
      $ 627 "Case 7"
      $ 628 "TM_St_Completin≔get_time(STATE_Times[STATE-1])"
      global TM_St_Completin=get_time(STATE_Times[STATE-1])
    elif (8 == switch_1):
      $ 629 "Case 8"
      $ 630 "TM_St_Complete≔get_time(STATE_Times[STATE-1])"
      global TM_St_Complete=get_time(STATE_Times[STATE-1])
    elif (9 == switch_1):
      $ 631 "Case 9"
      $ 632 "TM_St_Holding≔get_time(STATE_Times[STATE-1])"
      global TM_St_Holding=get_time(STATE_Times[STATE-1])
    elif (10 == switch_1):
      $ 633 "Case 10"
      $ 634 "TM_St_Held≔get_time(STATE_Times[STATE-1])"
      global TM_St_Held=get_time(STATE_Times[STATE-1])
    elif (11 == switch_1):
      $ 635 "Case 11"
      $ 636 "TM_St_Unholding≔get_time(STATE_Times[STATE-1])"
      global TM_St_Unholding=get_time(STATE_Times[STATE-1])
    elif (12 == switch_1):
      $ 637 "Case 12"
      $ 638 "TM_St_Suspendin≔get_time(STATE_Times[STATE-1])"
      global TM_St_Suspendin=get_time(STATE_Times[STATE-1])
    elif (13 == switch_1):
      $ 639 "Case 13"
      $ 640 "TM_St_Suspended≔get_time(STATE_Times[STATE-1])"
      global TM_St_Suspended=get_time(STATE_Times[STATE-1])
    elif (14 == switch_1):
      $ 641 "Case 14"
      $ 642 "TM_St_Unsuspend≔get_time(STATE_Times[STATE-1])"
      global TM_St_Unsuspend=get_time(STATE_Times[STATE-1])
    elif (15 == switch_1):
      $ 643 "Case 15"
      $ 644 "TM_St_Aborting≔get_time(STATE_Times[STATE-1])"
      global TM_St_Aborting=get_time(STATE_Times[STATE-1])
    elif (16 == switch_1):
      $ 645 "Case 16"
      $ 646 "TM_St_Aborted≔get_time(STATE_Times[STATE-1])"
      global TM_St_Aborted=get_time(STATE_Times[STATE-1])
    elif (17 == switch_1):
      $ 647 "Case 17"
      $ 648 "TM_St_Clearing≔get_time(STATE_Times[STATE-1])"
      global TM_St_Clearing=get_time(STATE_Times[STATE-1])
    end
    $ 650 "Wait: 0.1"
    sleep(0.1)
  end
end
